Fanuc KAREL source: KA00180.KL

PROGRAM KA00180
%NOLOCKGROUP
VAR
  SRC: ARRAY[4] OF STRING[20]
  DST: ARRAY[4] OF JOINTPOS
BEGIN
  DST = SRC
END KA00180
